(* PLC project Ejercicio_Tanque.project, CODESYS CODESYS V3.5 SP22 Patch 3 *)
(* stored: creationDateTime 2026-11-02T23:05:42.3674008, modificationDateTime 2026-10-01T10:32:36.9707997 *)

PROGRAM PLC_PRG

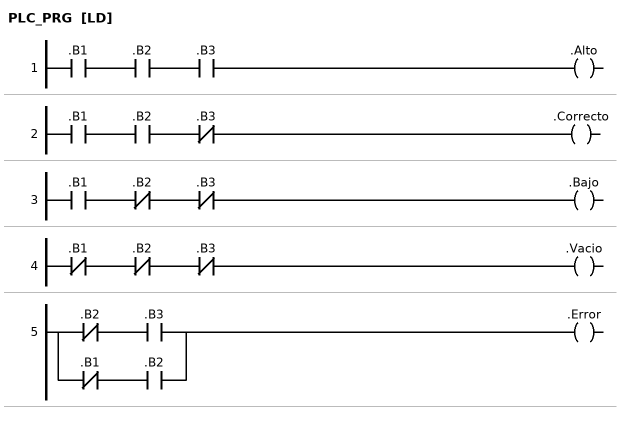
(* LD diagram, written out as Structured Text *)
(* Nivel de llenado muy alto (overflow) *)

.Alto := .B1 AND .B2 AND .B3;
(* Nivel de llenado correcto *)

.Correcto := .B1 AND .B2 AND NOT .B3;
(* Nivel de llenado muy bajo *)

.Bajo := .B1 AND NOT .B2 AND NOT .B3;
(* Nivel del tanque vacío *)

.Vacio := NOT .B1 AND NOT .B2 AND NOT .B3;
(* Casos de Error *)

.Error := NOT .B2 AND .B3 OR NOT .B1 AND .B2;
END_PROGRAM

CONFIGURATION Device
  RESOURCE Application ON PLC
    VAR_GLOBAL  (* GVL *)
      B1 : BOOL;  (* Sensor 1 (Vacío) *)
      B2 : BOOL;  (* Sensor 2 (Normal) *)
      B3 : BOOL;  (* Sensor 3 (OverFlow) *)
      Alto : BOOL;  (* H3 Nivel muy alto *)
      Correcto : BOOL;  (* H1 Nivel Correcto *)
      Bajo : BOOL;  (* H2 Nivel muy bajo *)
      Vacio : BOOL;  (* H4 Nivel Vacío *)
      Error : BOOL;  (* H5 Error *)
    END_VAR
    TASK MainTask(INTERVAL := T#20ms, PRIORITY := 1);
    TASK VISU_TASK(INTERVAL := T#100ms, PRIORITY := 31);
    PROGRAM PLC_PRG WITH MainTask : PLC_PRG;
    PROGRAM VisuElems.Visu_Prg WITH VISU_TASK : VisuElems.Visu_Prg;
  END_RESOURCE
END_CONFIGURATION
